Fanuc KAREL source: NC0063.KL

PROGRAM NC0063
%NOLOCKGROUP
ROUTINE R
VAR
  X : INTEGER
  I1 : INTEGER
  I2 : INTEGER
BEGIN
  X = 1
  FOR I1 = 1 TO 2 DO
    FOR I2 = 1 TO 2 DO
      X = X + 1
    ENDFOR
  ENDFOR
END R
BEGIN
  R
END NC0063
